(* IEC 61131-3 sources: SafePLC-Gen-Evaluation/Evaluation Results/dexpi/run_01, 2 files *)

(* ---- io_declarations.st ---- *)
(* ==================================================  *)
(* PLC I/O Variable Declarations — CODESYS 3.5  *)
(* Generated by SafePLC-Gen Multimodal  *)
(* ==================================================  *)

VAR_GLOBAL
    (* --- Analog Inputs ---  *)
    PI_4712.01_Raw               AT %IW0       : INT := 0;    (* PI-4712.01 — Pressure indicator (local gauge) on line  *)
    PICSA_4712.02_Raw            AT %IW2       : INT := 0;    (* PICSA-4712.02 — Pressure indicating controller with safe  *)
    TICSA_4750.03_Raw            AT %IW4       : INT := 0;    (* TICSA-4750.03 — Temperature indicating controller with s  *)
    (* --- Analog Outputs ---  *)
    PVA_4712.02_Out              AT %QW0       : INT := 0;    (* PVA-4712.02 — Pressure control valve (PVA - pressure v  *)
    TV_4750.03_Out               AT %QW2       : INT := 0;    (* TV-4750.03 — Temperature control valve on utility (he  *)
    (* --- Digital Inputs ---  *)
    HS_4750.01                   AT %IX0.0     : BOOL := FALSE;    (* HS-4750.01 — Hand switch / selector switch (HS) locat  *)
    (* --- Digital Outputs ---  *)
    XV_MNc_47124                 AT %QX0.0     : BOOL := FALSE;    (* XV-MNc-47124 — Check valve (non-return) on line MNc 471  *)
END_VAR

(* ---- generated_code.st ---- *)
(* Generated by SafePLC-Gen Multimodal — CODESYS 3.5 *)
(* IEC 61131-3 Structured Text *)
(* Date: 2026-04-25T13:33:38.376272 *)

PROGRAM PLC_Control

VAR
    TICSA_4750_03_Raw            AT %IW4       : INT := 0;
    PICSA_4712_02_Raw            AT %IW2       : INT := 0;
    PI_4712_01_Raw               AT %IW0       : INT := 0;
    PVA_4712_02_Out              AT %QW0       : INT := 0;
    TV_4750_03_Out               AT %QW2       : INT := 0;
    HS_4750_01                   AT %IX0.0     : BOOL := FALSE;
    XV_MNc_47124                 AT %QX0.0     : BOOL := FALSE;
    ESTOP                        AT %IX0.1     : BOOL := FALSE;
    MANUAL_RESET                 AT %IX0.2     : BOOL := FALSE;
END_VAR

VAR
    TICSA_4750_03_Scaled         : REAL := 0.0;
    PICSA_4712_02_Scaled         : REAL := 0.0;
    PI_4712_01_Scaled            : REAL := 0.0;

    TICSA_4750_03_HH_SP          : REAL := 180.0;
    TICSA_4750_03_H_SP           : REAL := 160.0;
    TICSA_4750_03_L_SP           : REAL := 20.0;
    TICSA_4750_03_LL_SP          : REAL := 10.0;
    TICSA_4750_03_Deadband       : REAL := 2.0;

    PICSA_4712_02_HH_SP          : REAL := 90.0;
    PICSA_4712_02_H_SP           : REAL := 80.0;
    PICSA_4712_02_L_SP           : REAL := 10.0;
    PICSA_4712_02_LL_SP          : REAL := 5.0;
    PICSA_4712_02_Deadband       : REAL := 1.0;

    PI_4712_01_HH_SP             : REAL := 90.0;
    PI_4712_01_H_SP              : REAL := 80.0;
    PI_4712_01_L_SP              : REAL := 10.0;
    PI_4712_01_LL_SP             : REAL := 5.0;
    PI_4712_01_Deadband          : REAL := 1.0;

    TICSA_4750_03_H              : BOOL := FALSE;
    TICSA_4750_03_L              : BOOL := FALSE;
    TICSA_4750_03_HH_Set         : BOOL := FALSE;
    TICSA_4750_03_HH_Rst         : BOOL := FALSE;
    TICSA_4750_03_LL_Set         : BOOL := FALSE;
    TICSA_4750_03_LL_Rst         : BOOL := FALSE;
    TICSA_4750_03_HH_Latch       : SR := (S1 := FALSE, R := FALSE);
    TICSA_4750_03_LL_Latch       : SR := (S1 := FALSE, R := FALSE);
    TICSA_4750_03_HH_Ack         : BOOL := FALSE;
    TICSA_4750_03_LL_Ack         : BOOL := FALSE;

    PICSA_4712_02_H              : BOOL := FALSE;
    PICSA_4712_02_L              : BOOL := FALSE;
    PICSA_4712_02_HH_Set         : BOOL := FALSE;
    PICSA_4712_02_HH_Rst         : BOOL := FALSE;
    PICSA_4712_02_LL_Set         : BOOL := FALSE;
    PICSA_4712_02_LL_Rst         : BOOL := FALSE;
    PICSA_4712_02_HH_Latch       : SR := (S1 := FALSE, R := FALSE);
    PICSA_4712_02_LL_Latch       : SR := (S1 := FALSE, R := FALSE);
    PICSA_4712_02_HH_Ack         : BOOL := FALSE;
    PICSA_4712_02_LL_Ack         : BOOL := FALSE;

    PI_4712_01_H                 : BOOL := FALSE;
    PI_4712_01_L                 : BOOL := FALSE;
    PI_4712_01_HH_Set            : BOOL := FALSE;
    PI_4712_01_HH_Rst            : BOOL := FALSE;
    PI_4712_01_LL_Set            : BOOL := FALSE;
    PI_4712_01_LL_Rst            : BOOL := FALSE;
    PI_4712_01_HH_Latch          : SR := (S1 := FALSE, R := FALSE);
    PI_4712_01_LL_Latch          : SR := (S1 := FALSE, R := FALSE);
    PI_4712_01_HH_Ack            : BOOL := FALSE;
    PI_4712_01_LL_Ack            : BOOL := FALSE;

    LOOP_4750_03_TRIP            : BOOL := FALSE;
    LOOP_4712_02_TRIP            : BOOL := FALSE;
    LOOP_104_01_TRIP             : BOOL := FALSE;
    TICSA_4750_03_HH             : BOOL := FALSE;
    TICSA_4750_03_LL             : BOOL := FALSE;
    PICSA_4712_02_HH             : BOOL := FALSE;
    PICSA_4712_02_LL             : BOOL := FALSE;
    SV_104_01_HH                 : BOOL := FALSE;
    SV_104_01_LL                 : BOOL := FALSE;
    SAFE_STATE                   : BOOL := FALSE;

    TICSA_4750_03_SP             : REAL := 80.0;
    TICSA_4750_03_Error          : REAL := 0.0;
    TICSA_4750_03_Integral       : REAL := 0.0;
    TICSA_4750_03_Kp             : REAL := 1.5;
    TICSA_4750_03_Ki             : REAL := 0.05;
    TICSA_4750_03_Output_Pct     : REAL := 0.0;

    PICSA_4712_02_SP             : REAL := 50.0;
    PICSA_4712_02_Error          : REAL := 0.0;
    PICSA_4712_02_Integral       : REAL := 0.0;
    PICSA_4712_02_Kp             : REAL := 1.2;
    PICSA_4712_02_Ki             : REAL := 0.04;
    PICSA_4712_02_Output_Pct     : REAL := 0.0;

    SV_104_01_Out                : BOOL := FALSE;
    HV_H_1007_N3_Out             : BOOL := FALSE;
    HV_H_1007_N4_Out             : BOOL := FALSE;
    HV_HS_4750_FC_Out            : BOOL := FALSE;
    HV_73KH12_25_inlet_Out       : BOOL := FALSE;
    HV_73KH12_25_outlet_Out      : BOOL := FALSE;
    HV_73KH12_bypass_Out         : BOOL := FALSE;
    HV_MNc_47126_block_Out       : BOOL := FALSE;
    HV_Q_80_block_Out            : BOOL := FALSE;

    System_Alarm                 : BOOL := FALSE;
    FirstScan                    : BOOL := TRUE;
END_VAR

IF FirstScan THEN
    LOOP_4750_03_TRIP        := TRUE;
    LOOP_4712_02_TRIP        := TRUE;
    LOOP_104_01_TRIP         := TRUE;
    SAFE_STATE               := TRUE;
    TV_4750_03_Out           := 6554;
    PVA_4712_02_Out          := 6554;
    XV_MNc_47124             := FALSE;
    SV_104_01_Out            := FALSE;
    HV_H_1007_N3_Out         := FALSE;
    HV_H_1007_N4_Out         := FALSE;
    HV_HS_4750_FC_Out        := FALSE;
    HV_73KH12_25_inlet_Out   := FALSE;
    HV_73KH12_25_outlet_Out  := FALSE;
    HV_73KH12_bypass_Out     := FALSE;
    HV_MNc_47126_block_Out   := FALSE;
    HV_Q_80_block_Out        := FALSE;
    TICSA_4750_03_HH_Latch(S1 := FALSE, R := TRUE);
    TICSA_4750_03_LL_Latch(S1 := FALSE, R := TRUE);
    PICSA_4712_02_HH_Latch(S1 := FALSE, R := TRUE);
    PICSA_4712_02_LL_Latch(S1 := FALSE, R := TRUE);
    PI_4712_01_HH_Latch(S1 := FALSE, R := TRUE);
    PI_4712_01_LL_Latch(S1 := FALSE, R := TRUE);
    FirstScan                := FALSE;
    RETURN;
END_IF;

TICSA_4750_03_Scaled := ((INT_TO_REAL(TICSA_4750_03_Raw) - 6554.0) / (32767.0 - 6554.0)) * 200.0;
PICSA_4712_02_Scaled := ((INT_TO_REAL(PICSA_4712_02_Raw) - 6554.0) / (32767.0 - 6554.0)) * 100.0;
PI_4712_01_Scaled    := ((INT_TO_REAL(PI_4712_01_Raw)    - 6554.0) / (32767.0 - 6554.0)) * 100.0;

TICSA_4750_03_HH := TICSA_4750_03_Scaled >= TICSA_4750_03_HH_SP;
TICSA_4750_03_LL := TICSA_4750_03_Scaled <= TICSA_4750_03_LL_SP;
PICSA_4712_02_HH := PICSA_4712_02_Scaled >= PICSA_4712_02_HH_SP;
PICSA_4712_02_LL := PICSA_4712_02_Scaled <= PICSA_4712_02_LL_SP;

IF TICSA_4750_03_HH OR TICSA_4750_03_LL THEN
    LOOP_4750_03_TRIP := TRUE;
ELSIF LOOP_4750_03_TRIP AND MANUAL_RESET AND NOT TICSA_4750_03_HH AND NOT TICSA_4750_03_LL THEN
    LOOP_4750_03_TRIP := FALSE;
END_IF;

IF PICSA_4712_02_HH OR PICSA_4712_02_LL THEN
    LOOP_4712_02_TRIP := TRUE;
ELSIF LOOP_4712_02_TRIP AND MANUAL_RESET AND NOT PICSA_4712_02_HH AND NOT PICSA_4712_02_LL THEN
    LOOP_4712_02_TRIP := FALSE;
END_IF;

IF SV_104_01_HH OR SV_104_01_LL THEN
    LOOP_104_01_TRIP := TRUE;
ELSIF LOOP_104_01_TRIP AND MANUAL_RESET AND NOT SV_104_01_HH AND NOT SV_104_01_LL THEN
    LOOP_104_01_TRIP := FALSE;
END_IF;

SAFE_STATE := ESTOP OR LOOP_4750_03_TRIP OR LOOP_4712_02_TRIP OR LOOP_104_01_TRIP;

IF NOT SAFE_STATE THEN
    TICSA_4750_03_Error    := TICSA_4750_03_SP - TICSA_4750_03_Scaled;
    TICSA_4750_03_Integral := TICSA_4750_03_Integral + (TICSA_4750_03_Ki * TICSA_4750_03_Error);
    IF TICSA_4750_03_Integral > 100.0 THEN
        TICSA_4750_03_Integral := 100.0;
    ELSIF TICSA_4750_03_Integral < 0.0 THEN
        TICSA_4750_03_Integral := 0.0;
    END_IF;
    TICSA_4750_03_Output_Pct := (TICSA_4750_03_Kp * TICSA_4750_03_Error) + TICSA_4750_03_Integral;
    IF TICSA_4750_03_Output_Pct > 100.0 THEN
        TICSA_4750_03_Output_Pct := 100.0;
    ELSIF TICSA_4750_03_Output_Pct < 0.0 THEN
        TICSA_4750_03_Output_Pct := 0.0;
    END_IF;
    TV_4750_03_Out := REAL_TO_INT(6554.0 + (TICSA_4750_03_Output_Pct / 100.0) * (32767.0 - 6554.0));
ELSE
    TV_4750_03_Out := 6554;
END_IF;

IF NOT SAFE_STATE THEN
    PICSA_4712_02_Error    := PICSA_4712_02_SP - PICSA_4712_02_Scaled;
    PICSA_4712_02_Integral := PICSA_4712_02_Integral + (PICSA_4712_02_Ki * PICSA_4712_02_Error);
    IF PICSA_4712_02_Integral > 100.0 THEN
        PICSA_4712_02_Integral := 100.0;
    ELSIF PICSA_4712_02_Integral < 0.0 THEN
        PICSA_4712_02_Integral := 0.0;
    END_IF;
    PICSA_4712_02_Output_Pct := (PICSA_4712_02_Kp * PICSA_4712_02_Error) + PICSA_4712_02_Integral;
    IF PICSA_4712_02_Output_Pct > 100.0 THEN
        PICSA_4712_02_Output_Pct := 100.0;
    ELSIF PICSA_4712_02_Output_Pct < 0.0 THEN
        PICSA_4712_02_Output_Pct := 0.0;
    END_IF;
    PVA_4712_02_Out := REAL_TO_INT(6554.0 + (PICSA_4712_02_Output_Pct / 100.0) * (32767.0 - 6554.0));
ELSE
    PVA_4712_02_Out := 6554;
END_IF;

IF NOT SAFE_STATE THEN
    XV_MNc_47124             := HS_4750_01;
    SV_104_01_Out            := TRUE;
    HV_H_1007_N3_Out         := TRUE;
    HV_H_1007_N4_Out         := TRUE;
    HV_HS_4750_FC_Out        := HS_4750_01;
    HV_73KH12_25_inlet_Out   := TRUE;
    HV_73KH12_25_outlet_Out  := TRUE;
    HV_73KH12_bypass_Out     := FALSE;
    HV_MNc_47126_block_Out   := TRUE;
    HV_Q_80_block_Out        := TRUE;
ELSE
    XV_MNc_47124             := FALSE;
    SV_104_01_Out            := FALSE;
    HV_H_1007_N3_Out         := FALSE;
    HV_H_1007_N4_Out         := FALSE;
    HV_HS_4750_FC_Out        := FALSE;
    HV_73KH12_25_inlet_Out   := FALSE;
    HV_73KH12_25_outlet_Out  := FALSE;
    HV_73KH12_bypass_Out     := FALSE;
    HV_MNc_47126_block_Out   := FALSE;
    HV_Q_80_block_Out        := FALSE;
END_IF;

IF TICSA_4750_03_Scaled >= TICSA_4750_03_HH_SP THEN
    TICSA_4750_03_HH_Set := TRUE;
ELSIF TICSA_4750_03_Scaled <= (TICSA_4750_03_HH_SP - TICSA_4750_03_Deadband) THEN
    TICSA_4750_03_HH_Set := FALSE;
END_IF;
TICSA_4750_03_HH_Rst := TICSA_4750_03_HH_Ack AND NOT TICSA_4750_03_HH_Set;
TICSA_4750_03_HH_Latch(S1 := TICSA_4750_03_HH_Set, R := TICSA_4750_03_HH_Rst);

IF TICSA_4750_03_Scaled <= TICSA_4750_03_LL_SP THEN
    TICSA_4750_03_LL_Set := TRUE;
ELSIF TICSA_4750_03_Scaled >= (TICSA_4750_03_LL_SP + TICSA_4750_03_Deadband) THEN
    TICSA_4750_03_LL_Set := FALSE;
END_IF;
TICSA_4750_03_LL_Rst := TICSA_4750_03_LL_Ack AND NOT TICSA_4750_03_LL_Set;
TICSA_4750_03_LL_Latch(S1 := TICSA_4750_03_LL_Set, R := TICSA_4750_03_LL_Rst);

TICSA_4750_03_H := TICSA_4750_03_Scaled >= TICSA_4750_03_H_SP;
TICSA_4750_03_L := TICSA_4750_03_Scaled <= TICSA_4750_03_L_SP;

IF PICSA_4712_02_Scaled >= PICSA_4712_02_HH_SP THEN
    PICSA_4712_02_HH_Set := TRUE;
ELSIF PICSA_4712_02_Scaled <= (PICSA_4712_02_HH_SP - PICSA_4712_02_Deadband) THEN
    PICSA_4712_02_HH_Set := FALSE;
END_IF;
PICSA_4712_02_HH_Rst := PICSA_4712_02_HH_Ack AND NOT PICSA_4712_02_HH_Set;
PICSA_4712_02_HH_Latch(S1 := PICSA_4712_02_HH_Set, R := PICSA_4712_02_HH_Rst);

IF PICSA_4712_02_Scaled <= PICSA_4712_02_LL_SP THEN
    PICSA_4712_02_LL_Set := TRUE;
ELSIF PICSA_4712_02_Scaled >= (PICSA_4712_02_LL_SP + PICSA_4712_02_Deadband) THEN
    PICSA_4712_02_LL_Set := FALSE;
END_IF;
PICSA_4712_02_LL_Rst := PICSA_4712_02_LL_Ack AND NOT PICSA_4712_02_LL_Set;
PICSA_4712_02_LL_Latch(S1 := PICSA_4712_02_LL_Set, R := PICSA_4712_02_LL_Rst);

PICSA_4712_02_H := PICSA_4712_02_Scaled >= PICSA_4712_02_H_SP;
PICSA_4712_02_L := PICSA_4712_02_Scaled <= PICSA_4712_02_L_SP;

IF PI_4712_01_Scaled >= PI_4712_01_HH_SP THEN
    PI_4712_01_HH_Set := TRUE;
ELSIF PI_4712_01_Scaled <= (PI_4712_01_HH_SP - PI_4712_01_Deadband) THEN
    PI_4712_01_HH_Set := FALSE;
END_IF;
PI_4712_01_HH_Rst := PI_4712_01_HH_Ack AND NOT PI_4712_01_HH_Set;
PI_4712_01_HH_Latch(S1 := PI_4712_01_HH_Set, R := PI_4712_01_HH_Rst);

IF PI_4712_01_Scaled <= PI_4712_01_LL_SP THEN
    PI_4712_01_LL_Set := TRUE;
ELSIF PI_4712_01_Scaled >= (PI_4712_01_LL_SP + PI_4712_01_Deadband) THEN
    PI_4712_01_LL_Set := FALSE;
END_IF;
PI_4712_01_LL_Rst := PI_4712_01_LL_Ack AND NOT PI_4712_01_LL_Set;
PI_4712_01_LL_Latch(S1 := PI_4712_01_LL_Set, R := PI_4712_01_LL_Rst);

PI_4712_01_H := PI_4712_01_Scaled >= PI_4712_01_H_SP;
PI_4712_01_L := PI_4712_01_Scaled <= PI_4712_01_L_SP;

System_Alarm :=
    TICSA_4750_03_HH_Latch.Q1 OR TICSA_4750_03_LL_Latch.Q1 OR
    TICSA_4750_03_H            OR TICSA_4750_03_L            OR
    PICSA_4712_02_HH_Latch.Q1 OR PICSA_4712_02_LL_Latch.Q1 OR
    PICSA_4712_02_H            OR PICSA_4712_02_L            OR
    PI_4712_01_HH_Latch.Q1    OR PI_4712_01_LL_Latch.Q1    OR
    PI_4712_01_H               OR PI_4712_01_L               OR
    SAFE_STATE;

END_PROGRAM
